(* IEC 61131-3 sources: traffic-lights/PLC_TrafficLights/Class/SafetyBaseFSoE (part 2) *)

  if WriteDOsUsed then
    for i := 0 to WriteDOsUsed-1 do
      SetDORunState(Handle:=aWritePDOs[i].Handle, NewState:=_BUS_IF_RUN_STATE_CONT_RUN);
    end_for;
  end_if;

  if usAnalogInputReadDOsUsed then
    for i := 0 to usAnalogInputReadDOsUsed-1 do
      SetDORunState(Handle:=aAnalogInputReadDOs[i].Handle, NewState:=_BUS_IF_RUN_STATE_CONT_RUN);
    end_for;
  end_if;

  if ReadFastUnsafeDOsUsed then
    for i := 0 to ReadFastUnsafeDOsUsed-1 do
      SetDORunState(Handle:=aFastUnsafeReadDOs[i].Handle, NewState:=_BUS_IF_RUN_STATE_CONT_RUN);
    end_for;
  end_if;

  if WriteFastUnsafeDOsUsed then
    for i := 0 to WriteFastUnsafeDOsUsed-1 do
      SetDORunState(Handle:=aFastUnsafeWriteDOs[i].Handle, NewState:=_BUS_IF_RUN_STATE_CONT_RUN);
    end_for;
  end_if;

END_FUNCTION

FUNCTION VIRTUAL SafetyBaseFSoE::StopDO
  VAR
    i : USINT;
  END_VAR

  // disable the DOs
  SetDORunState(Handle:=TempReadDO.Handle, NewState:=_BUS_IF_RUN_STATE_NO_RUN);

  SetDORunState(Handle:=TempWriteDO.Handle, NewState:=_BUS_IF_RUN_STATE_NO_RUN);

  if ReadDOsUsed then
    for i := 0 to ReadDOsUsed-1 do
      SetDORunState(Handle:=aReadPDOs[i].Handle, NewState:=_BUS_IF_RUN_STATE_NO_RUN);
    end_for;
  end_if;

  if WriteDOsUsed then
    for i := 0 to WriteDOsUsed-1 do
      SetDORunState(Handle:=aWritePDOs[i].Handle, NewState:=_BUS_IF_RUN_STATE_NO_RUN);
    end_for;
  end_if;

  if usAnalogInputReadDOsUsed then
    for i := 0 to usAnalogInputReadDOsUsed-1 do
      SetDORunState(Handle:=aAnalogInputReadDOs[i].Handle, NewState:=_BUS_IF_RUN_STATE_NO_RUN);
    end_for;
  end_if;

  if ReadFastUnsafeDOsUsed then
    for i := 0 to ReadFastUnsafeDOsUsed-1 do
      SetDORunState(Handle:=aFastUnsafeReadDOs[i].Handle, NewState:=_BUS_IF_RUN_STATE_NO_RUN);
    end_for;
  end_if;

  if WriteFastUnsafeDOsUsed then
    for i := 0 to WriteFastUnsafeDOsUsed-1 do
      SetDORunState(Handle:=aFastUnsafeWriteDOs[i].Handle, NewState:=_BUS_IF_RUN_STATE_NO_RUN);
    end_for;
  end_if;

END_FUNCTION

FUNCTION VIRTUAL SafetyBaseFSoE::InitBuffers
  VAR_OUTPUT
    sd_retval 	: DINT;
  END_VAR

  sd_retval := -1;

  //allocate memory for outgoing SDO (one SDO possible)
  p_SDOOutputBuffer$^void := ToStdLib.Malloc(size := SBF_SDO_MAX_LENGTH);

  if ( p_SDOOutputBuffer = NIL ) then
    SetSafetyState(NewState:=_MemAllocFailed);
    return;
  end_if;

  //allocate memory for incoming SDO list (number of SDO is dynamical)
  //following elements will be added dynamical

  //allocate list
  InputBufferAllocatedNo := SBF_SDO_BUFFER_ALLOC_BLOCK;
  p_SDOInputBuffer$^void := ToStdLib.Malloc(size := InputBufferAllocatedNo * SBF_SDO_MAX_LENGTH);

  if ( p_SDOInputBuffer = NIL ) then
    SetSafetyState(NewState:=_MemAllocFailed);
    return;
  end_if;

  //all buffers initialized
  sd_retval := 0;

END_FUNCTION

FUNCTION VIRTUAL SafetyBaseFSoE::GetSafetyNumber
  VAR_OUTPUT
    sd_retval 	: DINT;
  END_VAR
  VAR
    TempPathInfo  : PathInfoType;
    MyPara 	  : CmdStruct;
    MyResult	: results;
  END_VAR

  sd_retval := SDOStdRequ ( us_Command      := SBF_SDO_COMMAND_GET_SAFENBR
                          , p_us_RespData   := ( #SafetyNumber )$^USINT
                          , us_RespLength   := sizeof(SafetyNumber)
                          );

  if ( sd_retval <> 0 ) then
    if b_NoSafetyLogged = FALSE then
      b_NoSafetyLogged := TRUE;
      LogError("@01D8 (SafetyBaseFSoE::GetSafetyNumber) [SL] No Safety Number available!");
    end_if;
  elsif pConfigMem then
    // store safety number in config memory
    pConfigMem^$HDINT := SafetyNumber;
  end_if;

  sd_retval := SDOStdRequ ( us_Command      := SBF_SDO_COMMAND_GET_FW_VERSION
                          , p_us_RespData   := ( #sFirmwareVersion )$^USINT
                          , us_RespLength   := sizeof(FirmwareVersionType)
                          );

  if ( sd_retval = 0 ) then
    FirmwareVersion := sFirmwareVersion.RevMinor OR (sFirmwareVersion.RevMajor SHL 16);

    // Minor Versions starting with 9xxx mark Bootloader versions
    if (sFirmwareVersion.RevMinor >= 9000) & (sFirmwareVersion.RevMinor < 10000) then
      LogError("@01D9 (SafetyBaseFSoE::GetSafetyNumber) Bootloader version of safety firmware detected! Download a firmware or contact Sigmatek Support!");
    end_if;

    //Minor Versions higher than 338 mark versions which support the readout of the safety retry counters.
    if (sFirmwareVersion.RevMinor >= SBF_RETRY_COUNTER_AVAILABLE_MINOR_REV) & (sFirmwareVersion.RevMajor = SBF_RETRY_COUNTER_AVAILABLE_MAJOR_REV) then
      b_RetryCounterAvailable := TRUE;
    else
      b_RetryCounterAvailable := FALSE;
      //Call Method to set retrycounter servers of safety modules to -1
      SetRetryCounter();
    end_if;
  else
    SetSafetyState(NewState:=_ReadFWVerFailed);
    LogError("@01DA (SafetyBaseFSoE::GetSafetyNumber) No Firmware Version available!");
  end_if;

  InitPathInfo(#TempPathInfo);

  // add own safety number to routing table
  sd_retval := AddRoutingElement( ud_SafeNumber       := SafetyNumber
                                , ud_thisp            := this$UDINT
                                , pObject             := #TempPathInfo
                                );

  // give the manager more details about the module
  if pSafetyManagerThis then
    MyPara.uiCmd := CMD_SM_ADD_MODULE_INFO;
    MyPara.aPara[0] := THIS$DINT;
    MyPara.aPara[1] := SafetyNumber$DINT;
    MyPara.aPara[2] := FirmwareVersion$DINT;
    MyPara.aPara[3] := 16#FF; // fake FPGA_Version (only needed for CDIAS CPUs)
    MyPara.aPara[4] := to_DINT(p_ObjectPath^$USINT) + 1; // size of path (length + 1 for the length information)
    MyPara.aPara[5] := p_ObjectPath$DINT;
    pSafetyManagerThis^.NewInst(#MyPara, #MyResult);
  else
    LogError("@01DB (SafetyBaseFSoE::GetSafetyNumber) Couldn't find object of HwControl class, which is needed for safety time synchronisation!");
  end_if;

END_FUNCTION

FUNCTION SafetyBaseFSoE::SafetyBaseFSoE
  VAR_OUTPUT
    ret_code 	: ConfStates;
  END_VAR

#ifdef HWC_LogInit
  HWC_LogInit();
#endif

  //get interface for safety functions
  if ( OS_CILGET(INTERFACE_SAFETY, #pISafety)) then
    pISafety := NIL;

    LogError("@01DC (SafetyBaseFSoE::SafetyBaseFSoE) No Safety Interface found!");
  end_if;

  // initialize it with FALSE, if there is anything on local CDIAS it will change to TRUE
  b_SafetyOnLocalCDIAS := FALSE;

  // initialize module count with 0
  ModuleSyncNo := 0;

  ret_code := C_OK;

END_FUNCTION

#pragma warning(disable:0073);
FUNCTION VIRTUAL SafetyBaseFSoE::UpDateNotStd
  VAR_INPUT
    calloption 	: UDINT;
  END_VAR

END_FUNCTION
#pragma warning(default:0073);

FUNCTION VIRTUAL SafetyBaseFSoE::ReadSDOConfig
  VAR_INPUT
    p_SDORequestBuffer 	: ^SafetyBaseFSoE::SDORequReadConfig;
    p_SDOResponseBuffer 	: ^SafetyBaseFSoE::SDORespReadConfig;
    pModule 	: ^SafetyBaseFSoE::PathInfoType;
    pListHeader 	: ^SafetyBaseFSoE::PathInfoType;
  END_VAR
  VAR_OUTPUT
    sd_retval 	: DINT;
  END_VAR
  VAR
    ud_Address                    : UDINT;
    ud_ListLength_Address         : UDINT;
    ud_ListLength                 : UDINT;
    ud_TmpCnt                     : UDINT;
    i                             : UDINT;
    ud_ModulePathLen_Max          : UDINT;
    ud_ModulePathCompLen_Max      : UDINT;
    ud_ListHeaderPathLen_Max      : UDINT;
    ud_ListHeaderPathCompLen_Max  : UDINT;
    us_DataLength_Max             : USINT;
    ud_ListBaseAddress            : UDINT;
    ud_ListAddressMax             : UDINT;
    ud_CntUnsafeOutputs           : UDINT;
    ud_CntUnsafeInputs            : UDINT;
    ud_ActAddress                 : UDINT;  // actual offset in application memory (where to find the values in run mode)
    ud_UnsafeBDINT_Offset         : UDINT;  // actual offset in application memory (where to find the unsafe variables in run mode)
    ud_ActBlockType               : UDINT;
    ud_TmpAddress                 : UDINT;
    ud_TmpStrLen                  : UDINT;
    p_TmpBlockedData              : ^void;
    ud_ActStrLen                  : UDINT;
    us_BlockedTransferLength      : USINT;
    BoolOuts                      : UDINT;
    DintOuts                      : UDINT;
    TempModuleConfig              : t_ModuleCfg;
    pChar                         : ^CHAR;
    TempPath                      : ARRAY [0..99] OF USINT;
    PathOfThisCPU                 : ARRAY [0..99] OF USINT;
    GotOwnPath                    : BOOL;
    TempPdoConfig                 : t_PdoCfg;
    pBitMasks                     : ^BDINT;
    ActBitMask                    : BDINT;
    ud_skipLength                 : UDINT; //++pr
    b_CfgTypeV2                   : BOOL; // FALSE means there is no support of new time synchronisation/new general purpose register
    TmpCRC                        : HDINT;
    ud_ContainerBlockType         : UDINT;
    b_CfgTypeV3                   : BOOL;
    ud_ConfigLength               : UDINT;
    hd_DynParaVersion             : UDINT;
    DynamicParameterHeader        : t_DynamicParameterHeader;
    b_IsFSoE                      : BOOL;
    DynHeadSize                   : UDINT;
    AddressServiceDataSize        : UDINT;
    b_IprCodeLengthAvailable      : BOOL;  //TRUE, SCP211 is used
    ud_CntFastUnsafeOutputs       : UDINT;
    ud_CntFastUnsafeInputs        : UDINT;
    ud_FastUnsafe_Offset_In       : UDINT; // actual offset in application memory (where to find the unsafe variables in run mode)
    ud_FastUnsafe_Offset_Out      : UDINT; // actual offset in application memory (where to find the unsafe variables in run mode)
    ud_TmpLength                  : UDINT;

  END_VAR

  //minimum length of path: 2 bytes length, 1 byte domain info, 1 byte bus type and 1 byte port  => we use maximum so we don't have dynamic memory => don't fragment heap
  ud_ModulePathLen_Max          := 128;
  ud_ModulePathCompLen_Max      := 128;
  ud_ListHeaderPathLen_Max      := 128;
  ud_ListHeaderPathCompLen_Max  := 128;

  NewConfigType := ConfigState_NotInitialized;

  // reset flags before checking the config
  sFlexCon.FoundNodeInConfig := FALSE;
  sFlexCon.FoundHostInConfig := FALSE;
  b_IprCodeLengthAvailable        := FALSE;

  // also reset the servers
  if sFlexCon.pCommand & sFlexCon.pStateMachine & sFlexCon.pHostSafetyNumber then
    sFlexCon.pCommand^          := 0;
    sFlexCon.pStateMachine^     := 0;
    sFlexCon.pHostSafetyNumber^ := 0;
  end_if;

  //initialize header-data for request

  //calculate length without crc
  p_SDORequestBuffer^.StdHeader.Len := sizeof(SDORequReadConfig) - sizeof(SDOHeader.StdHeader.CRC);

  //type
  p_SDORequestBuffer^.StdHeader.Typ := SDO_STD;

  //command for reading config data
  p_SDORequestBuffer^.StdHeader.Cmd := SBF_SDO_COMMAND_READ;

  //read crc of whole config data

  //send request and receive data
  sd_retval := SDOReadCfgRequ ( p_SDORequestBuffer  := p_SDORequestBuffer
                              , p_SDOResponseBuffer := p_SDOResponseBuffer
                              , ud_Address          := SBF_SDO_ADDRESS_CONFIG_DATA + SBF_SDO_OFFSET_CONFIG_CRC_ALL
                              , us_Length           := 4
                              );

  //no response
  if ( sd_retval <> 0 ) then
    LogError("@01DD (SafetyBaseFSoE::ReadSDOConfig) Error reading CRC of config data.");
    return;
  end_if;

  // save crc and remember the time
  DesignerPrjConfigCRC := p_SDOResponseBuffer^.ud_Data;
  ud_LastCrcCheck := ops.tAbsolute;
  b_CheckCRC := TRUE;

  //read length of whole config data

  //send request and receive data
  sd_retval := SDOReadCfgRequ ( p_SDORequestBuffer  := p_SDORequestBuffer
                              , p_SDOResponseBuffer := p_SDOResponseBuffer
                              , ud_Address          := SBF_SDO_ADDRESS_CONFIG_DATA + SBF_SDO_OFFSET_CONFIG_LEN_ALL
                              , us_Length           := 4
                              );

  //no response
  if ( sd_retval <> 0 ) then
    LogError("@01DE (SafetyBaseFSoE::ReadSDOConfig) Error reading length of config data.");
    return;
  end_if;

  //no config data available
  if ( p_SDOResponseBuffer^.ud_Data = 16#FFFF_FFFF ) then
    LogError("@01DF (SafetyBaseFSoE::ReadSDOConfig) No config data available..");
    b_ReadConfigFailed := TRUE;
    return;
  end_if;

  ud_ConfigLength := p_SDOResponseBuffer^.ud_Data;

  // get BlockType
  //send request and receive data
  sd_retval := SDOReadCfgRequ ( p_SDORequestBuffer  := p_SDORequestBuffer
                              , p_SDOResponseBuffer := p_SDOResponseBuffer
                              , ud_Address          := SBF_SDO_ADDRESS_CONFIG_DATA + SBF_SDO_OFFSET_CONFIG_BLOCKTYPE
                              , us_Length           := 4
                              );
  //no response, error
  if ( sd_retval <> 0 ) then
    LogError("@01E0 (SafetyBaseFSoE::ReadSDOConfig) Error getting the block type of the header.");
    return;
  end_if;

  ud_ContainerBlockType := p_SDOResponseBuffer^.ud_Data;

  // check if it's a new version of the configuration
  if (ud_ContainerBlockType = SBF_BLKTYPE_CFG_CONTAINER_V3)       |
     (ud_ContainerBlockType = SBF_BLKTYPE_CFG_CONTAINER_V3_SLAVE)     |
     (ud_ContainerBlockType = SBF_BLKTYPE_CFG_CONTAINER_V3_SLAVE_OPTIONAL) then

    //read dynamic header length (how many data are attached to the header)

    //send request and receive data
    sd_retval := SDOReadCfgRequ ( p_SDORequestBuffer  := p_SDORequestBuffer
                                , p_SDOResponseBuffer := p_SDOResponseBuffer
                                , ud_Address          := SBF_SDO_ADDRESS_CONFIG_DATA + SBF_SDO_OFFSET_CONFIG_LEN_HEAD
                                , us_Length           := 4
                                );

    //no response
    if ( sd_retval <> 0 ) then
      LogError("@01E1 (SafetyBaseFSoE::ReadSDOConfig) Error reading length of dynamic header data.");
      return;
    end_if;

    // plausibility check for data length
    if p_SDOResponseBuffer^.ud_Data > 1000 then
      sd_retval := -1;
      LogError("@01E2 (SafetyBaseFSoE::ReadSDOConfig) Invalid length of dynamic header data.");
      return;
    end_if;

    // the length info contains: size of length info + size of time info + size of additional data

    //start address of first list: address of dynamic length + length according to length info
    ud_ListBaseAddress := SBF_SDO_ADDRESS_CONFIG_DATA + SBF_SDO_OFFSET_CONFIG_LEN_HEAD + p_SDOResponseBuffer^.ud_Data;

    DynHeadSize := p_SDOResponseBuffer^.ud_Data;

    // if we got at least 4 byte additional header data, it's the version of the dynamic parameters => read it
    if DynHeadSize >= 12 then
      //send request and receive data
      sd_retval := SDOReadCfgRequ ( p_SDORequestBuffer  := p_SDORequestBuffer
                                  , p_SDOResponseBuffer := p_SDOResponseBuffer
                                  , ud_Address          := SBF_SDO_ADDRESS_CONFIG_DATA + SBF_SDO_OFFSET_CONFIG_LEN_HEAD + 8
                                  , us_Length           := 4
                                  );

      //no response
      if ( sd_retval <> 0 ) then
        LogError("@01E3 (SafetyBaseFSoE::ReadSDOConfig) Error reading version of dynamic header data.");
        return;
      end_if;

      hd_DynParaVersion := p_SDOResponseBuffer^.ud_Data;
    else
      LogError("@01E4 (SafetyBaseFSoE::ReadSDOConfig) Data structure error in config! No bytes for the dynamic parameter version (according to length info).");
      return;
    end_if;

    // if we got at least 8 byte additional header data, the next 4 bytes are the flags => read it
    if DynHeadSize >= 16 then
      //send request and receive data
      sd_retval := SDOReadCfgRequ ( p_SDORequestBuffer  := p_SDORequestBuffer
                                  , p_SDOResponseBuffer := p_SDOResponseBuffer
                                  , ud_Address          := SBF_SDO_ADDRESS_CONFIG_DATA + SBF_SDO_OFFSET_CONFIG_LEN_HEAD + 12
                                  , us_Length           := 4
                                  );

      //no response
      if ( sd_retval <> 0 ) then
        LogError("@023D (SafetyBaseFSoE::ReadSDOConfig) Error reading flags of dynamic header data.");
        return;
      end_if;

      b_IsFSoE := (p_SDOResponseBuffer^.ud_Data AND 1) <> 0;

      // if we got the FSoE bit set => read the FSoE config
      if b_IsFSoE then
        GetFSoEConnectionInfos(p_SDORequestBuffer   := p_SDORequestBuffer
                             , p_SDOResponseBuffer  := p_SDOResponseBuffer
                             );
      end_if;

      if DynHeadSize >= 20 then
        //send request and receive data
        sd_retval := SDOReadCfgRequ ( p_SDORequestBuffer  := p_SDORequestBuffer
                                    , p_SDOResponseBuffer := p_SDOResponseBuffer
                                    , ud_Address          := SBF_SDO_ADDRESS_CONFIG_DATA + SBF_SDO_OFFSET_CONFIG_LEN_HEAD + 16
                                    , us_Length           := 4
                                    );

        //no response
        if ( sd_retval <> 0 ) then
          LogError("@023D (SafetyBaseFSoE::ReadSDOConfig) Error reading flags of dynamic header data.");
          return;
        end_if;

        b_IprCodeLengthAvailable := (p_SDOResponseBuffer^.ud_Data AND 1) <> 0;

        // if there are fast unsafe variables to read
        if uiPDOReadSizeFastUnsafeVar then

          //malloc FastUnsafe Output Buffer
          pFastUnsafeOutBuffer := ToStdLib.Malloc(size:=uiPDOReadSizeFastUnsafeVar);

          if pFastUnsafeOutBuffer = NIL then
            LogError("@0784 (SafetyBaseFSoE::ReadSDOConfig) Failed to allocate memory for outputbuffer.");
            return;
          else
            // init buffer
            _memset(dest:=pFastUnsafeOutBuffer, usByte:=0x00, cntr:=uiPDOReadSizeFastUnsafeVar);
          end_if;
        end_if;

        // if there are fast unsafe variables to write
        if uiPDOWriteSizeFastUnsafeVar then

          //malloc FastUnsafe Input Buffer
          pFastUnsafeInBuffer := ToStdLib.Malloc(size:=uiPDOWriteSizeFastUnsafeVar);

          if pFastUnsafeInBuffer = NIL then
            LogError("@0785 (SafetyBaseFSoE::ReadSDOConfig) Failed to allocate memory for inputbuffer.");
            return;
          else
            // init buffer
            _memset(dest:=pFastUnsafeInBuffer, usByte:=0x00, cntr:=uiPDOWriteSizeFastUnsafeVar);
          end_if;
        end_if;
      end_if;

    else
      LogError("@01E4 (SafetyBaseFSoE::ReadSDOConfig) Data structure error in config! No bytes for the dynamic parameter version (according to length info).");
      return;
    end_if;
  else
    // old version => no dynamic header, the first list starts where the dynamic header length would be

    //start address of first list: address of time info + size of time info
    ud_ListBaseAddress := SBF_SDO_ADDRESS_CONFIG_DATA + SBF_SDO_OFFSET_CONFIG_LEN_HEAD + sizeof(UDINT);
  end_if;

  GotOwnPath := FALSE;

  //highest address for config data
  ud_ListAddressMax := SDO_ADDRESS_CONFIG_DATA + SDO_OFFSET_CONFIG_LEN_ALL + ud_ConfigLength;

  //max. length of data to read with one request
  us_DataLength_Max := SBF_SDO_MAX_LENGTH - sizeof(SDORespReadConfig) + sizeof(SDORespReadConfig.ud_Data);

  while ( ud_ListBaseAddress < ud_ListAddressMax ) do

    //first read length of path in list-header

    //read path in list-header
    sd_retval := ReadModulePath ( p_SDORequestBuffer          := p_SDORequestBuffer
                                , p_SDOResponseBuffer         := p_SDOResponseBuffer
                                , p_ud_Address                := #ud_ListBaseAddress
                                , pModule                     := pListHeader
                                , p_ud_ModulePathLen_Max      := #ud_ListHeaderPathLen_Max
                                , p_ud_ModulePathCompLen_Max  := #ud_ListHeaderPathCompLen_Max
                                , us_SDOMaxDataSize           := us_DataLength_Max
                                );

    //no response, error
    if ( sd_retval <> 0 ) then
      LogError("@01E5 (SafetyBaseFSoE::ReadSDOConfig) Error reading module path out of config data.");
      return;
    end_if;

    // remember our own uncompressed path (first listheader path in the memory)
    if pListHeader^.p_us_Path & (GotOwnPath = FALSE) then
      GotOwnPath := TRUE;

      // remember the path
      _memcpy(ptr1:=#PathOfThisCPU[0], ptr2:=pListHeader^.p_us_Path, cntr:=(pListHeader^.p_us_Path$^UINT)^ + 2);
    end_if;

    //read length of download data in list-header (=LengthOverall) and save address
    //to calculate later the address of next list-header
    //address = last address + 4 byte (CRC)
    ud_ListLength_Address := ud_ListBaseAddress + 4;

    //send request and receive data
    sd_retval := SDOReadCfgRequ ( p_SDORequestBuffer  := p_SDORequestBuffer
                                , p_SDOResponseBuffer := p_SDOResponseBuffer
                                , ud_Address          := ud_ListLength_Address
                                , us_Length           := 4
                                );

    //no response
    if ( sd_retval <> 0 ) then
      LogError("@01E6 (SafetyBaseFSoE::ReadSDOConfig) Failed to read out the length of the download data within the configuration.");
      return;
    end_if;

    //save length of list
    ud_ListLength := p_SDOResponseBuffer^.ud_Data;

    //                                                   v
    //address of LengthOverall + 4 bytes (LengthOverall, BlockType, ModuleID)
    ud_Address := ud_ListLength_Address + 4;

    // get BlockType
    //send request and receive data
    sd_retval := SDOReadCfgRequ ( p_SDORequestBuffer  := p_SDORequestBuffer
                                , p_SDOResponseBuffer := p_SDOResponseBuffer
                                , ud_Address          := ud_Address
                                , us_Length           := 4
                                );
    //no response, error
    if ( sd_retval <> 0 ) then
      LogError("@01E7 (SafetyBaseFSoE::ReadSDOConfig) Error getting the block type.");
      return;
    end_if;

    ud_ActBlockType := p_SDOResponseBuffer^.ud_Data;

    case ud_ActBlockType of
//**********************************************************************************************************************************************************
      SBF_BLKTYPE_CFG_CPU,
      SBF_BLKTYPE_CFG_CPU_OPTIONAL , // if we don't need data from an external cpu
      SBF_BLKTYPE_CFG_MASTER_CPU:
        //add other CPUs to routing table

        // if there is a valid module path
        if pListHeader^.p_us_Path <> NIL then
          //add module to routing tabs
          sd_retval := AddModuleToRoutingTabs ( pModule       := pListHeader
                                              , pListHeader   := pListHeader
                                              , b_IsOptional  := (ud_ActBlockType = SBF_BLKTYPE_CFG_CPU_OPTIONAL)
                                              );

          if (sd_retval <> 0 ) then
            if ( SafetyState <> _ModFromCfgNotFound ) then
              LogError("@01E8 (SafetyBaseFSoE::ReadSDOConfig) Failed to add cpu module to routing tabs.");
              return;
            end_if;
          end_if;

          TempModuleConfig.Info := 0;
          TempModuleConfig.DestCRCNo := 0;
          TempModuleConfig.pDestCRCs := NIL;
          TempModuleConfig.PdoOutLen := 0;

          TempModuleConfig.Info.IsOptional  := (ud_ActBlockType = SBF_BLKTYPE_CFG_CPU_OPTIONAL);
          TempModuleConfig.InterfaceCRC     := 0;

          // Remember the path (uncompressed and compressed)
          TempModuleConfig.PathLen := pListHeader^.p_us_Path^$UINT + 2;
          TempModuleConfig.pPath := pListHeader^.p_us_Path;

          TempModuleConfig.CompPathLen := pListHeader^.ui_PathCompLen;
          TempModuleConfig.pCompPath := pListHeader^.p_us_PathComp;

          // if it's our own path, remember the safety number
          if (PathOfThisCPU[0]$UINT = (pListHeader^.p_us_Path$^UINT)^) & (ToStdLib.MemCmp(#PathOfThisCPU[0], pListHeader^.p_us_Path, PathOfThisCPU[0]$UINT + 2) = 0) then
            TempModuleConfig.SafetyNbr := SafetyNumber;
            //safe config of scp modul (own path)
            SafeActModuleConfig(TempModuleConfig);
          else
            TempModuleConfig.SafetyNbr := 0;
          end_if;

          // only when there is a manager
          if pSafetyManagerThis then
            AddModuleToCfg(TempModuleConfig);
          end_if;
        end_if;

//**********************************************************************************************************************************************************
      SBF_BLKTYPE_CFG_SLAVE_COMPR,
      SBF_BLKTYPE_CFG_SLAVE_COMPR_OPTIONAL: //Blocktyp der über die komprimierte Gesamtkonfiguration einer Slave-CPU gegeben wird
        //add other CPUs to routing table

        // if there is a valid module path
        if pListHeader^.p_us_Path <> NIL then
          //add module to routing tabs
          sd_retval := AddModuleToRoutingTabs ( pModule       := pListHeader
                                              , pListHeader   := pListHeader
                                              , b_IsOptional  := (ud_ActBlockType = SBF_BLKTYPE_CFG_SLAVE_COMPR_OPTIONAL)
                                              );

          if (sd_retval <> 0 ) then
            if ( SafetyState <> _ModFromCfgNotFound ) then
              LogError("@0270 (SafetyBaseFSoE::ReadSDOConfig) Slave: Failed to add cpu module to routing tabs.");
              return;
            end_if;
          end_if;

          // we skip the config till we get to the interface information of this slave (if it's the source of an interface frame we have to remember it)

          //address of LengthOverall + 3 * 4 bytes (LengthOverall, BlockType, ModuleID) => now the address points to FUB offset
          ud_Address := ud_ListLength_Address + 12;

          //skip FUB offset
          ud_Address += 4;

          // get no of FUB´s
          //send request and receive data
          sd_retval := SDOReadCfgRequ ( p_SDORequestBuffer  := p_SDORequestBuffer
                                      , p_SDOResponseBuffer := p_SDOResponseBuffer
                                      , ud_Address          := ud_Address
                                      , us_Length           := 4
                                      );
          //no response, error
          if ( sd_retval <> 0 ) then
            LogError("@01E9 (SafetyBaseFSoE::ReadSDOConfig) Slave: Error getting the FUB number.");
            return;
          end_if;

          ud_TmpCnt := p_SDOResponseBuffer^.ud_Data;

          // skip no of FUB´s and FUB´s
          ud_Address += (4 + (ud_TmpCnt * 4));

          // get length of path
          //send request and receive data
          sd_retval := SDOReadCfgRequ ( p_SDORequestBuffer  := p_SDORequestBuffer
                                      , p_SDOResponseBuffer := p_SDOResponseBuffer
                                      , ud_Address          := ud_Address
                                      , us_Length           := 4
                                      );
          //no response, error
          if ( sd_retval <> 0 ) then
            LogError("@01EA (SafetyBaseFSoE::ReadSDOConfig) Slave: Error getting the path length.");
            return;
          end_if;

          ud_TmpCnt := p_SDOResponseBuffer^.ud_Data;

          // skip length of path and the path
          ud_Address += (4 + ud_TmpCnt);

          // get length of comp path
          //send request and receive data
          sd_retval := SDOReadCfgRequ ( p_SDORequestBuffer  := p_SDORequestBuffer
                                      , p_SDOResponseBuffer := p_SDOResponseBuffer
                                      , ud_Address          := ud_Address
                                      , us_Length           := 4
                                      );
          //no response, error
          if ( sd_retval <> 0 ) then
            LogError("@01EB (SafetyBaseFSoE::ReadSDOConfig) Slave: Error getting the comp path length.");
            return;
          end_if;

          ud_TmpCnt := p_SDOResponseBuffer^.ud_Data;

          // skip length of comp path and the comp path
          ud_Address += (4 + ud_TmpCnt);

          // skip CRC and LengthOverall to get to the Blocktyp (Modul-Downloaddaten)
          ud_Address += 8;

          // get the block type
          //send request and receive data
          sd_retval := SDOReadCfgRequ ( p_SDORequestBuffer  := p_SDORequestBuffer
                                      , p_SDOResponseBuffer := p_SDOResponseBuffer
                                      , ud_Address          := ud_Address
                                      , us_Length           := 4
                                      );
          //no response, error
          if ( sd_retval <> 0 ) then
            LogError("@01EC (SafetyBaseFSoE::ReadSDOConfig) Slave: Error getting the block type of a slave config.");
            return;
          end_if;

          ud_TmpCnt := p_SDOResponseBuffer^.ud_Data;

          // check if it's a new version of the configuration
          if (ud_TmpCnt = SBF_BLKTYPE_CFG_CONTAINER_V3)       |
             (ud_TmpCnt = SBF_BLKTYPE_CFG_CONTAINER_V3_SLAVE)     |
             (ud_TmpCnt = SBF_BLKTYPE_CFG_CONTAINER_V3_SLAVE_OPTIONAL) then

            // skip blocktype to get to the dynamic header length (how many data are attached to the header)
            ud_Address += 4;

            //send request and receive data
            sd_retval := SDOReadCfgRequ ( p_SDORequestBuffer  := p_SDORequestBuffer
                                        , p_SDOResponseBuffer := p_SDOResponseBuffer
                                        , ud_Address          := ud_Address
                                        , us_Length           := 4
                                        );

            //no response
            if ( sd_retval <> 0 ) then
              LogError("@01ED (SafetyBaseFSoE::ReadSDOConfig) Error reading length of dynamic header data of a slave config.");
              return;
            end_if;

            // plausibility check for data length
            if p_SDOResponseBuffer^.ud_Data > 1000 then
              sd_retval := -1;
              LogError("@01EE (SafetyBaseFSoE::ReadSDOConfig) Invalid length of dynamic header data of a slave config.");
              return;
            end_if;

            // the length info contains: size of length info + size of time info + size of additional data

            // skip the additional data to get to the path length
            ud_Address += p_SDOResponseBuffer^.ud_Data;
          else
            // old version => no dynamic header, so we skip only blocktype and time info
            ud_Address += 8;
          end_if;

          // get the path length
          //send request and receive data
          sd_retval := SDOReadCfgRequ ( p_SDORequestBuffer  := p_SDORequestBuffer
                                      , p_SDOResponseBuffer := p_SDOResponseBuffer
                                      , ud_Address          := ud_Address
                                      , us_Length           := 4
                                      );
          //no response, error
          if ( sd_retval <> 0 ) then
            LogError("@01EA (SafetyBaseFSoE::ReadSDOConfig) Slave: Error getting the path length.");
            return;
          end_if;

          ud_TmpCnt := p_SDOResponseBuffer^.ud_Data;

          // skip length of path and the path
          ud_Address += (4 + ud_TmpCnt);

          // get length of comp path
          //send request and receive data
          sd_retval := SDOReadCfgRequ ( p_SDORequestBuffer  := p_SDORequestBuffer
                                      , p_SDOResponseBuffer := p_SDOResponseBuffer
                                      , ud_Address          := ud_Address
                                      , us_Length           := 4
                                      );
          //no response, error
          if ( sd_retval <> 0 ) then
            LogError("@01EB (SafetyBaseFSoE::ReadSDOConfig) Slave: Error getting the comp path length.");
            return;
          end_if;

          ud_TmpCnt := p_SDOResponseBuffer^.ud_Data;

          // skip length of comp path and the comp path
          ud_Address += (4 + ud_TmpCnt);

          // skip CRC, LengthOverall, Blocktyp (Modul-Downloaddaten), ModuleID
          ud_Address += 16;

          // get the InterfaceCRC
          //send request and receive data
          sd_retval := SDOReadCfgRequ ( p_SDORequestBuffer  := p_SDORequestBuffer
                                      , p_SDOResponseBuffer := p_SDOResponseBuffer
                                      , ud_Address          := ud_Address
                                      , us_Length           := 4
                                      );
          //no response, error
          if ( sd_retval <> 0 ) then
            LogError("@01EF (SafetyBaseFSoE::ReadSDOConfig) Slave: Error getting the Inteface-CRC.");
            return;
          end_if;

          TmpCRC := p_SDOResponseBuffer^.ud_Data;

          //add slave information to config
          AddSlaveToCfg ( pModule       := pListHeader
                        , b_IsOptional  := (ud_ActBlockType = SBF_BLKTYPE_CFG_SLAVE_COMPR_OPTIONAL)
                        , b_IsInterface := (TmpCRC <> 0)
                        , InterfaceCRC  := TmpCRC
                        );

        end_if;

//**********************************************************************************************************************************************************
      SBF_BLKTYPE_CFG_REV: // revision

        // check if the list is long enough for a String (more bytes than just the header)
        if ud_ListLength > 12 then

          //address of LengthOverall + 3 * 4 bytes (LengthOverall, BlockType, ModuleID) => now the address points to the revision string
          ud_Address := ud_ListLength_Address + 12;

          //read out the string (length = LengthOverall - length header)

          // get memory for the string
          if pPrjNameStr = NIL then
            PrjNameMemLen := ud_ListLength$USINT - 12;
            pPrjNameStr$^void := ToStdLib.Malloc(size := PrjNameMemLen + 1);
          else
            if PrjNameMemLen <> (ud_ListLength$USINT - 12) then
              PrjNameMemLen := ud_ListLength$USINT - 12;
              pPrjNameStr$^void := ToStdLib.ReAlloc(mptr:=pPrjNameStr, newsize:=PrjNameMemLen + 1);
            end_if;
          end_if;

          // check if we got a memory
          if pPrjNameStr then

            _memset(dest:=pPrjNameStr, usByte:=0, cntr:=PrjNameMemLen+1);

            ud_ActStrLen := ud_TmpStrLen := PrjNameMemLen;
            ud_TmpAddress := ud_Address;

            IF p_BlockedTransferMemory = NIL THEN
              sd_retval := -100;
              SetSafetyState(NewState:=_MemAllocFailed);
              RETURN;
            END_IF;

            IF ud_BlockedTransferMemorySize < (ud_TmpStrLen + 1) THEN
              p_BlockedTransferMemory := ToStdLib.ReAlloc(mptr:=p_BlockedTransferMemory, newsize:=GetNewMemSize(ud_TmpStrLen + 1));
              IF p_BlockedTransferMemory = NIL THEN
                ud_BlockedTransferMemorySize := 0;
                sd_retval := -100;
                SetSafetyState(NewState:=_MemAllocFailed);
                RETURN;
              ELSE
                ud_BlockedTransferMemorySize := GetNewMemSize(ud_TmpStrLen + 1);
              END_IF;
            END_IF;

            ToStdLib.MemSet(dest:=p_BlockedTransferMemory, value:=0, size:=ud_BlockedTransferMemorySize);

            p_TmpBlockedData := p_BlockedTransferMemory;

            us_BlockedTransferLength := BlockedTransferLength(ud_Datalength:=ud_TmpStrLen, us_MaxBlocklength:=60);

            while us_BlockedTransferLength do

              // get name
              sd_retval := SDOReadCfgRequ ( p_SDORequestBuffer  := p_SDORequestBuffer
                                          , p_SDOResponseBuffer := p_SDOResponseBuffer
                                          , ud_Address          := ud_TmpAddress
                                          , us_Length           := us_BlockedTransferLength
                                          , b_UseCache          := us_BlockedTransferLength < us_DataLength_Max
                                          );
              //no response
              if ( sd_retval <> 0 ) then
                LogError("@01F0 (SafetyBaseFSoE::ReadSDOConfig) Reading Revision failed.");
                return;
              end_if;

              ToStdLib.MemCpy(dest:=p_TmpBlockedData,
                               source:=#p_SDOResponseBuffer^.ud_Data,
                               size:=us_BlockedTransferLength);

              p_TmpBlockedData += us_BlockedTransferLength;
              ud_TmpAddress += us_BlockedTransferLength;
              ud_TmpStrLen -= us_BlockedTransferLength;

              us_BlockedTransferLength := BlockedTransferLength(ud_Datalength:=ud_TmpStrLen, us_MaxBlocklength:=60);

            end_while;

            ToStdLib.MemCpy(dest:=pPrjNameStr,
                             source:=p_BlockedTransferMemory,
                             size:=PrjNameMemLen+1);

            b_GotNewRevision := TRUE;

            // string is formed by: project name {TAB} project revision   => search for the tab
            pPrjRevStr := pPrjNameStr; // initialize pointer, because maybe there is no content in the projectname
            pChar := pPrjNameStr;
            while pChar^ do
              // check for tab sign
              if pChar^ = 9 then
                // at the next character our revision starts
                pPrjRevStr := pChar + sizeof(CHAR);

                // we change the tab to a string termination
                pChar^ := 0;

                // save the length of the name and the length of the project revision
                PrjNameStrLen := pChar$UDINT - pPrjNameStr$UDINT;
                PrjRevStrLen := PrjNameMemLen - PrjNameStrLen - sizeof(CHAR);
                exit;
              end_if;

              pChar += sizeof(CHAR);
            end_while;

            ShowProjectRevision();
          end_if;
        end_if;

//**********************************************************************************************************************************************************
      SBF_BLKTYPE_CFG_CRC: // CRC from Safety Application and HW-Tree

        // check if the list is long enough for a String (more bytes than just the header)
        if ud_ListLength > 12 then

          //address of LengthOverall + 3 * 4 bytes (LengthOverall, BlockType, ModuleID) => now the address points to the CRC values
          ud_Address := ud_ListLength_Address + 12;

          //read out the CRCs (length = 2 * 4 bytes)

          //send request and receive data
          sd_retval := SDOReadCfgRequ ( p_SDORequestBuffer  := p_SDORequestBuffer
                                      , p_SDOResponseBuffer := p_SDOResponseBuffer
                                      , ud_Address          := ud_Address
                                      , us_Length           := 2*sizeof(HDINT)
                                      );

          //no response
          if ( sd_retval <> 0 ) then
            LogError("@0797 (SafetyBaseFSoE::ReadSDOConfig) Reading CRC info of the safety designer project failed.");
            return;
          end_if;

          CRCInfo := p_SDOResponseBuffer^.ud_Data$t_CRCInfo;

          ApplCRC := CRCInfo.ApplCRC;
          HwCRC   := CRCInfo.HwCRC;
        end_if;

//**********************************************************************************************************************************************************
      SBF_BLKTYPE_CFG_INTERFACE,
      SBF_BLKTYPE_CFG_INTERFACE_OPTIONAL: // interface frame

        TempPdoConfig.Info := 0;

        //address of LengthOverall + 3 * 4 bytes (LengthOverall, BlockType, Module ID) => points to interface CRC
        ud_Address := ud_ListLength_Address + 12;

//*****************************************************************************
//**   INTERFACE CRC                                                         **
//*****************************************************************************

        //send request and receive data
        sd_retval := SDOReadCfgRequ ( p_SDORequestBuffer  := p_SDORequestBuffer
                                    , p_SDOResponseBuffer := p_SDOResponseBuffer
                                    , ud_Address          := ud_Address
                                    , us_Length           := 4
                                    );

        //no response
        if ( sd_retval <> 0 ) then
          LogError("@01F1 (SafetyBaseFSoE::ReadSDOConfig) Interface: Reading interface CRC of interface frame block failed.");
          return;
        end_if;

        TempPdoConfig.InterfaceCRC := p_SDOResponseBuffer^.ud_Data;

        // skip interface crc
        ud_Address += 4;

//*****************************************************************************
//**   LENGTH OF TOPOLOGY PATH OF INTERFACE FRAME                            **
//*****************************************************************************

        //send request and receive data
        sd_retval := SDOReadCfgRequ ( p_SDORequestBuffer  := p_SDORequestBuffer
                                    , p_SDOResponseBuffer := p_SDOResponseBuffer
                                    , ud_Address          := ud_Address
                                    , us_Length           := 4
                                    );

        //no response
        if ( sd_retval <> 0 ) then
          LogError("@01F2 (SafetyBaseFSoE::ReadSDOConfig) Interface: Reading length of topology path of interface frame block failed.");
          return;
        end_if;

        // skip path length
        ud_Address += 4;

        us_BlockedTransferLength := p_SDOResponseBuffer^.ud_Data$USINT;

//*****************************************************************************
//**   TOPOLOGY PATH OF INTERFACE FRAME                                      **
//*****************************************************************************

        //send request and receive data
        sd_retval := SDOReadCfgRequ ( p_SDORequestBuffer  := p_SDORequestBuffer
                                    , p_SDOResponseBuffer := p_SDOResponseBuffer
                                    , ud_Address          := ud_Address
                                    , us_Length           := us_BlockedTransferLength
                                    , b_UseCache          := us_BlockedTransferLength < us_DataLength_Max
                                    );

        //no response
        if ( sd_retval <> 0 ) then
          LogError("@01F3 (SafetyBaseFSoE::ReadSDOConfig) Interface: Reading topology path of interface frame block failed.");
          return;
        end_if;

        // remember the destination path
        _memcpy(ptr1:=#TempPath[0], ptr2:=#p_SDOResponseBuffer^.ud_Data, cntr:=us_BlockedTransferLength);

        // this is the source of the interface frame
        TempPdoConfig.SourcePathLen := TempPath[0]$UINT + 2;
        TempPdoConfig.pSourcePath   := #TempPath[0];

        // skip path
        ud_Address += us_BlockedTransferLength;

//*****************************************************************************
//**   LENGTH OF COMPRESSED TOPOLOGY PATH OF INTERFACE FRAME                 **
//*****************************************************************************

        //send request and receive data
        sd_retval := SDOReadCfgRequ ( p_SDORequestBuffer  := p_SDORequestBuffer
                                    , p_SDOResponseBuffer := p_SDOResponseBuffer
                                    , ud_Address          := ud_Address
                                    , us_Length           := 4
                                    );

        //no response
        if ( sd_retval <> 0 ) then
          LogError("@01F4 (SafetyBaseFSoE::ReadSDOConfig) Interface: Reading length of compressed topology path of interface frame block failed.");
          return;
        end_if;

        // skip path length
        ud_Address += 4;

        us_BlockedTransferLength := p_SDOResponseBuffer^.ud_Data$USINT;

//*****************************************************************************
//**   COMPRESSED TOPOLOGY PATH OF INTERFACE FRAME                           **
//*****************************************************************************

        //send request and receive data
        sd_retval := SDOReadCfgRequ ( p_SDORequestBuffer  := p_SDORequestBuffer
                                    , p_SDOResponseBuffer := p_SDOResponseBuffer
                                    , ud_Address          := ud_Address
                                    , us_Length           := us_BlockedTransferLength
                                    , b_UseCache          := us_BlockedTransferLength < us_DataLength_Max
                                    );

        //no response
        if ( sd_retval <> 0 ) then
          LogError("@01F5 (SafetyBaseFSoE::ReadSDOConfig) Interface: Reading compressed topology path of interface frame block failed.");
          return;
        end_if;

        // if it's an IP address => we need the compressed path for the source
        if p_SDOResponseBuffer^.ud_Data$USINT = 6 then
          // we may need this later (e.g. if it's an IP address)
          _memcpy(ptr1:=#TempPath[0], ptr2:=#p_SDOResponseBuffer^.ud_Data, cntr:=us_BlockedTransferLength);

          // this is the source of the interface frame
          TempPdoConfig.SourcePathLen := us_BlockedTransferLength;
          TempPdoConfig.Info.SrcPathIsCompressed := TRUE;

          if ((#p_SDOResponseBuffer^.ud_Data + 5)^$HDINT AND 16#00FFFFFF) = 0 then
            // special IP: (0.0.0.x)
            TempPdoConfig.Info.SrcPathIsCompressed := FALSE;  // Not valid IP
          end_if;
        end_if;

        // skip path and maximum cycle time
        ud_Address += us_BlockedTransferLength + 4;

  // here starts the data area (before we read only the list header

//*****************************************************************************
//**   INTERFACE CRC                                                         **
//*****************************************************************************

        //send request and receive data
        sd_retval := SDOReadCfgRequ ( p_SDORequestBuffer  := p_SDORequestBuffer
                                    , p_SDOResponseBuffer := p_SDOResponseBuffer
                                    , ud_Address          := ud_Address
                                    , us_Length           := 4
                                    );

        //no response
        if ( sd_retval <> 0 ) then
          LogError("@01F6 (SafetyBaseFSoE::ReadSDOConfig) Interface: Reading CRC of interface frame block failed.");
          return;
        end_if;

        TempPdoConfig.InterfaceCRC := p_SDOResponseBuffer^.ud_Data;

        // skip interface CRC
        ud_Address += 4;

//*****************************************************************************
//**   NUMBER OF BOOL INTERFACE VARIABLES IN THE PDO                         **
//*****************************************************************************

        //send request and receive data
        sd_retval := SDOReadCfgRequ ( p_SDORequestBuffer  := p_SDORequestBuffer
                                    , p_SDOResponseBuffer := p_SDOResponseBuffer
                                    , ud_Address          := ud_Address
                                    , us_Length           := 4
                                    );

        //no response
        if ( sd_retval <> 0 ) then
          LogError("@01F7 (SafetyBaseFSoE::ReadSDOConfig) Interface: Reading number of bool variables in the interface frame failed.");
          return;
        end_if;

        BoolOuts := p_SDOResponseBuffer^.ud_Data;

        // skip bool variables
        ud_Address += 4;

//*****************************************************************************
//**   NUMBER OF DINT INTERFACE VARIABLES IN THE PDO                         **
//*****************************************************************************

        //send request and receive data
        sd_retval := SDOReadCfgRequ ( p_SDORequestBuffer  := p_SDORequestBuffer
                                    , p_SDOResponseBuffer := p_SDOResponseBuffer
                                    , ud_Address          := ud_Address
                                    , us_Length           := 4
                                    );

        //no response
        if ( sd_retval <> 0 ) then
          LogError("@01F8 (SafetyBaseFSoE::ReadSDOConfig) Interface: Reading number of dint variables in the interface frame failed.");
          return;
        end_if;

        // skip dint variables
        ud_Address += 4;

        DintOuts := p_SDOResponseBuffer^.ud_Data;

        // if there are interface variables
        if BoolOuts | DintOuts then
          // calculate the length of the interface frame
          TempPdoConfig.PdoLen := CalcPDOLength(BoolOuts, DintOuts);

          // and the destination
          TempPdoConfig.DestPathLen   := PathOfThisCPU[0]$UINT + 2;
          TempPdoConfig.pDestPath     := #PathOfThisCPU[0];

          TempPdoConfig.Info.IsInterfacePDO := TRUE;
          TempPdoConfig.Info.IsOptional := (ud_ActBlockType = SBF_BLKTYPE_CFG_INTERFACE_OPTIONAL);

          // add the interface PDO to the list
          AddPdoToCfg(TempPdoConfig);
        else
          LogError("@01F9 (SafetyBaseFSoE::ReadSDOConfig) Interface: No interface variables found in interface blocktype.");
          return;
        end_if;

//**********************************************************************************************************************************************************
      SBF_BLKTYPE_CFG_MODULE_WITHOUT_CFG,
      SBF_BLKTYPE_CFG_MODULE_WITHOUT_CFG_OPT:      // module configurations
        TempModuleConfig.Info := 0;
        TempModuleConfig.DestCRCNo := 0;
        TempModuleConfig.pDestCRCs := NIL;
        case ud_ActBlockType of
          SBF_BLKTYPE_CFG_MODULE_WITHOUT_CFG_OPT:
            TempModuleConfig.Info.IsOptional := TRUE;
          else
            TempModuleConfig.Info.IsOptional := FALSE;
        end_case;

        BoolOuts := 0;
        DintOuts := 0;

        // Remember the path (uncompressed and compressed)
        TempModuleConfig.PathLen := pListHeader^.p_us_Path^$UINT + 2;
        TempModuleConfig.pPath := pListHeader^.p_us_Path;

        TempModuleConfig.CompPathLen := pListHeader^.ui_PathCompLen;
        TempModuleConfig.pCompPath := pListHeader^.p_us_PathComp;

        //add module to routing tabs
        sd_retval := AddModuleToRoutingTabs ( pModule       := pListHeader
                                            , pListHeader   := pListHeader
                                            , b_IsOptional  := TempModuleConfig.Info.IsOptional
                                            );

        if (sd_retval <> 0 ) then
          if ( SafetyState <> _ModFromCfgNotFound ) then
            LogError("@020D (SafetyBaseFSoE::ReadSDOConfig) Failed to add safe input module to routing tabs.");
            return;
          end_if;
        end_if;

//*****************************************************************************
//**   LIST HEADER                                                           **
//*****************************************************************************
//   Offset  Größe	Beschreibung
//    0x00	4 Byte	CRC32
//    0x04	4 Byte	Länge der Konfiguration (inkl. Längenfeld)
//    0x08	4 Byte	Block-Typ (nicht optional: 0x00000029; optional: 0x40000029)
//    0x0C	4 Byte	Modul-ID
//    0x10	4 Byte	Version der Konfiguration (0x00000000)
//*****************************************************************************

        //address of LengthOverall + 4 * 4 bytes (LengthOverall, BlockType, ModuleID, VersionConfig)
        ud_Address := ud_ListLength_Address + 16;

//*****************************************************************************
//    FSoE Konfiguration
//*****************************************************************************
//    0x14	4 Byte	Anzahl an FSoE-Verbindungen (0x00000001)
//*****************************************************************************
//    FSoE Konfiguration * Anzahl an FSoE-Verbindungen
//*****************************************************************************
//    0x18	4 Byte	Länge der FSoE-Konfiguration
//    0x1C	4 Byte	Flags (0x00000000)
//    0x20	2 Byte	Größe der sicheren Ausgänge in Byte
//    0x22	2 Byte	Größe der sicheren Eingänge in Byte
//    0x24	2 Byte	FSoE Slaveadresse
//    0x26	2 Byte	reserviert
//*****************************************************************************

        // skip entrys to read fsoe slave address
        ud_Address += 16;

        //send request and receive data
        sd_retval := SDOReadCfgRequ ( p_SDORequestBuffer  := p_SDORequestBuffer
                                    , p_SDOResponseBuffer := p_SDOResponseBuffer
                                    , ud_Address          := ud_Address
                                    , us_Length           := 4
                                    );

        //no response
        if ( sd_retval <> 0 ) then
          LogError("@01F6 (SafetyBaseFSoE::ReadSDOConfig) Reading interface CRC of interface frame block failed.");
          return;
        end_if;

        // only when there is a manager
        if pSafetyManagerThis then
          AddModuleToCfg(TempModuleConfig);
        end_if;

//**********************************************************************************************************************************************************
      SBF_BLKTYPE_CFG_MODULE,
      SBF_BLKTYPE_CFG_MODULE_V2,
      SBF_BLKTYPE_CFG_MODULE_OPTIONAL,
      SBF_BLKTYPE_CFG_CONTAINER_SLAVE,
      SBF_BLKTYPE_CFG_CONTAINER_SLAVE_OPTIONAL,
      SBF_BLKTYPE_CFG_MODULE_V3,
      SBF_BLKTYPE_CFG_MODULE_V3_OPTIONAL,
      SBF_BLKTYPE_CFG_CONTAINER_V3_SLAVE,
      SBF_BLKTYPE_CFG_CONTAINER_V3_SLAVE_OPTIONAL:      // module configurations
        TempModuleConfig.Info := 0;
        TempModuleConfig.DestCRCNo := 0;
        TempModuleConfig.pDestCRCs := NIL;
        case ud_ActBlockType of
          SBF_BLKTYPE_CFG_MODULE_OPTIONAL,
          SBF_BLKTYPE_CFG_CONTAINER_SLAVE_OPTIONAL,
          SBF_BLKTYPE_CFG_MODULE_V3_OPTIONAL,
          SBF_BLKTYPE_CFG_CONTAINER_V3_SLAVE_OPTIONAL:
            TempModuleConfig.Info.IsOptional := TRUE;
          else
            TempModuleConfig.Info.IsOptional := FALSE;
        end_case;

        b_CfgTypeV2 := (ud_ActBlockType <> SBF_BLKTYPE_CFG_MODULE);

        // check if it's a V3 config, because the structure of the IO List is different
        if (ud_ActBlockType = SBF_BLKTYPE_CFG_MODULE_V3) |
           (ud_ActBlockType = SBF_BLKTYPE_CFG_MODULE_V3_OPTIONAL) |
           (ud_ActBlockType = SBF_BLKTYPE_CFG_CONTAINER_V3_SLAVE) |
           (ud_ActBlockType = SBF_BLKTYPE_CFG_CONTAINER_V3_SLAVE_OPTIONAL) then
          b_CfgTypeV3 := TRUE;
        else
          b_CfgTypeV3 := FALSE;
        end_if;

        // if it's our own path, remember the type of module configuration
        if (PathOfThisCPU[0]$UINT = (pListHeader^.p_us_Path$^UINT)^) & (ToStdLib.MemCmp(#PathOfThisCPU[0], pListHeader^.p_us_Path, PathOfThisCPU[0]$UINT + 2) = 0) then
          // if config is already "old" dont change to "new". (can be set by block SBF_BLKTYPE_OLD_MODE_FLAG)
          if NewConfigType <> ConfigState_Old then
            NewConfigType := (b_CfgTypeV2$USINT + 1)$t_ConfigStateType;
          end_if;
        end_if;

        BoolOuts := 0;
        DintOuts := 0;

        // Remember the path (uncompressed and compressed)
        TempModuleConfig.PathLen := pListHeader^.p_us_Path^$UINT + 2;
        TempModuleConfig.pPath := pListHeader^.p_us_Path;

        TempModuleConfig.CompPathLen := pListHeader^.ui_PathCompLen;
        TempModuleConfig.pCompPath := pListHeader^.p_us_PathComp;

//*****************************************************************************
//**   LIST HEADER                                                           **
//*****************************************************************************

        //address of LengthOverall + 3 * 4 bytes (LengthOverall, BlockType, ModuleID)
        ud_Address := ud_ListLength_Address + 12;

        // only available at new modules
        if b_CfgTypeV2 then

//*****************************************************************************
//**   INTERFACE CRC                                                         **
//*****************************************************************************

          //send request and receive data
          sd_retval := SDOReadCfgRequ ( p_SDORequestBuffer  := p_SDORequestBuffer
                                      , p_SDOResponseBuffer := p_SDOResponseBuffer
                                      , ud_Address          := ud_Address
                                      , us_Length           := 4
                                      );

          //no response
          if ( sd_retval <> 0 ) then
            LogError("@01F6 (SafetyBaseFSoE::ReadSDOConfig) Reading interface CRC of interface frame block failed.");
            return;
          end_if;

          TempPdoConfig.InterfaceCRC := p_SDOResponseBuffer^.ud_Data;

          // skip interface crc
          ud_Address += 4;

//*****************************************************************************
//**   LENGTH OF TOPOLOGY PATH OF INTERFACE FRAME                            **
//*****************************************************************************

          //send request and receive data
          sd_retval := SDOReadCfgRequ ( p_SDORequestBuffer  := p_SDORequestBuffer
                                      , p_SDOResponseBuffer := p_SDOResponseBuffer
                                      , ud_Address          := ud_Address
                                      , us_Length           := 4
                                      );

          //no response
          if ( sd_retval <> 0 ) then
            LogError("@01F2 (SafetyBaseFSoE::ReadSDOConfig) Reading length of topology path of interface frame block failed.");
            return;
          end_if;

          // skip path length
          ud_Address += 4;

          us_BlockedTransferLength := p_SDOResponseBuffer^.ud_Data$USINT;

//*****************************************************************************
//**   TOPOLOGY PATH OF INTERFACE FRAME                                      **
//*****************************************************************************

          //send request and receive data
          sd_retval := SDOReadCfgRequ ( p_SDORequestBuffer  := p_SDORequestBuffer
                                      , p_SDOResponseBuffer := p_SDOResponseBuffer
                                      , ud_Address          := ud_Address
                                      , us_Length           := us_BlockedTransferLength
                                      , b_UseCache          := us_BlockedTransferLength < us_DataLength_Max
                                      );

          //no response
          if ( sd_retval <> 0 ) then
            LogError("@01F3 (SafetyBaseFSoE::ReadSDOConfig) Reading topology path of interface frame block failed.");
            return;
          end_if;

          // remember the destination path
          _memcpy(ptr1:=#TempPath[0], ptr2:=#p_SDOResponseBuffer^.ud_Data, cntr:=us_BlockedTransferLength);

          // skip path
          ud_Address += us_BlockedTransferLength;

//*****************************************************************************
//**   LENGTH OF COMPRESSED TOPOLOGY PATH OF INTERFACE FRAME                 **
//*****************************************************************************

          //send request and receive data
          sd_retval := SDOReadCfgRequ ( p_SDORequestBuffer  := p_SDORequestBuffer
                                      , p_SDOResponseBuffer := p_SDOResponseBuffer
                                      , ud_Address          := ud_Address
                                      , us_Length           := 4
                                      );

          //no response
          if ( sd_retval <> 0 ) then
            LogError("@01F4 (SafetyBaseFSoE::ReadSDOConfig) Reading length of compressed topology path of interface frame block failed.");
            return;
          end_if;

          // skip path length
          ud_Address += 4;

          us_BlockedTransferLength := p_SDOResponseBuffer^.ud_Data$USINT;

//*****************************************************************************
//**   COMPRESSED TOPOLOGY PATH OF INTERFACE FRAME                           **
//*****************************************************************************

          //send request and receive data
          sd_retval := SDOReadCfgRequ ( p_SDORequestBuffer  := p_SDORequestBuffer
                                      , p_SDOResponseBuffer := p_SDOResponseBuffer
                                      , ud_Address          := ud_Address
                                      , us_Length           := us_BlockedTransferLength
                                      , b_UseCache          := us_BlockedTransferLength < us_DataLength_Max
                                      );

          //no response
          if ( sd_retval <> 0 ) then
            LogError("@01F5 (SafetyBaseFSoE::ReadSDOConfig) Reading compressed topology path of interface frame block failed.");
            return;
          end_if;

          ud_Address += us_BlockedTransferLength;

          // skip max. cycle time
          ud_Address += 4;
        end_if;

        // on first 4 bytes is fix the system time
        ud_ActAddress := 4;

        // address in memory for unsafe BDINT variables
        ud_UnsafeBDINT_Offset := 0;

        // address on the module to access the fast unsafe variables via SDIAS (offset 1 for the message counter)
        ud_FastUnsafe_Offset_Out  := 1;
        ud_FastUnsafe_Offset_In   := 1;

//*****************************************************************************
//**   FSoE CONNECTION LIST                                                  **
//*****************************************************************************

        if b_IsFSoE then
          //send request and receive data
          sd_retval := SDOReadCfgRequ ( p_SDORequestBuffer  := p_SDORequestBuffer
                                      , p_SDOResponseBuffer := p_SDOResponseBuffer
                                      , ud_Address          := ud_Address
                                      , us_Length           := 4
                                      );

          //no response
          if ( sd_retval <> 0 ) then
            LogError("@0271 (SafetyBaseFSoE::ReadSDOConfig) Failed to get the number of FSoE elements.");
            return;
          end_if;

          ud_TmpCnt := p_SDOResponseBuffer^.ud_Data;

          // skip number of entries time
          ud_Address += 4;

          if ud_TmpCnt then
            for i := 1 to ud_TmpCnt do
              // read size of structure

              //send request and receive data
              sd_retval := SDOReadCfgRequ ( p_SDORequestBuffer  := p_SDORequestBuffer
                                          , p_SDOResponseBuffer := p_SDOResponseBuffer
                                          , ud_Address          := ud_Address
                                          , us_Length           := 4
                                          );

              //no response
              if ( sd_retval <> 0 ) then
                LogError("@0272 (SafetyBaseFSoE::ReadSDOConfig) Failed to read size of FSoE structure element.");
                return;
              end_if;

              // skip the whole entry since we got our info earlier via GetFSoEConnectionInfos()
              ud_Address += p_SDOResponseBuffer^.ud_Data;
            end_for;
          end_if;
        end_if;
(*

Aufbau Verbindungsliste:

Zuerst wird die Anzahl der Elemente in der Liste angegeben:

  ULONG nbrOfElements;                    // Anzahl der Elemente in der Liste

Danach kommen die einzelnen Listenelemente.
Der Anfang eines Listenelements ist auf 4 Byte ausgerichtet.

Aufbau des Listenelements:

  typedef struct FSOE_CONN_DSC
  {
    // Größe der Struktur (inkl. Längenfeld selbst)
    ULONG len;
    //! Flags
    //  Actually, type is 4 bytes in size but for compatibility reasons it is still used as 1 byte. As a result, bits 9-32 are currently not used.
    //  Bit1: 1, wenn FSoE-Master, 0=FSoE-Slave
    //  Bit2: 1, wenn die Slave-Adresse über den HW-Pfad ermittelt wird
    //  Bit3: 1, wenn CRC von der FW ermittelt werden muss
    //  Bit4: 1, wenn Interface und Slave
    //  Bit5: 1, wenn Multichannel verwendet werden, aber ein Multichannel ist nicht vorhanden und der Eingang auf 1 gesetzt wird.
    //  Bit6: 1, wenn der Adressvergabeservice verwendet werden soll
    //  Bit7: 1, wenn der Master beim Slave die Connection ID anfordert
    //  Bit8: 1, wenn es sich um ein HGW handelt
    //  Bit9: 1, wenn Assign Slave On Demand
    //  Bits 10-32: reserviert, sind auf 0 gesetzt und werden nicht ausgewertet
  #define FSOE_CONN_FLAGS_MASTER                    (1 << 0)
  #define FSOE_CONN_FLAGS_USE_HWPATH_AS_SLAVEADDR   (1 << 1)
    ULONG flags;
    //! Größe der sicheren Prozessdaten, die vom FSoE Master an den FSoE Slave übertragen werden
    // Wert kann nur 1 oder ein vielfaches von 2 sein (1, 2, 4, 6, ...)
    USHORT sizeSafeOutputs;
    //! Größe der sicheren Prozessdaten, die vom FSoE Slave an den FSoE Master übertragen werden
    // Wert kann nur 1 oder ein vielfaches von 2 sein (1, 2, 4, 6, ...)
    USHORT sizeSafeInputs;
    //! Safety over EtherCAT Slave Adresse der Safety over EtherCAT Connection
    // Bei einem Master ist das die Adresse des Ziels, bei einem Slave die eigene Adresse.
    // Wert 0 = Wert wird aus dem EEProm geholt oder über den HW-Pfad ermittelt
    // (HW-Pfad, wenn Flag FSOE_CONN_FLAGS_USE_HWPATH_AS_SLAVEADDR gesetzt ist)
    USHORT slaveAddress;

    // ==== die folgenden Daten gibt es nur im Master ====

    //! ConnectionId der Safety over EtherCAT Connection
    // Wert 0 = Wert wird aus dem EEProm geholt
    USHORT connectionId;

    //! Länge der Kommunikationsparameter, muss immer 2 sein
    USHORT commParaLength;
    //! FSoE Watchdog-Zeit in ms (nur für den Master relevant)
    USHORT watchdog_ms;
    //! Größe der Anwendungsparameter
    USHORT applParaLength;
    /*
----------------------------------------------------------------------
     * Bis hierher ist die Größe der Elemente in der Struktur fix.
     * Danach sind die Elemente mit variabler Größe angeordnet:
     *
     * Applikationsparameter:
     *    Die Applikationsparameter für ein SCP011 als FSoE Slave bestehen
     *    aus der Konfigurations-CRC (Listenheader) oder der Interface-CRC
     *    des Slaves.
     *
     * HW-Pfad: <-- ist auf 4 Byte ausgerichtet
     *    Wenn das Flag FSOE_CONN_FLAGS_USE_HWPATH_AS_SLAVEADDR gesetzt ist, dann
     *    ermittelt sich der Master die Adresse des Slaves anhand des hier
     *    angegebenen HW-Pfades.
     *    Wenn das Flag FSOE_CONN_FLAGS_USE_HWPATH_AS_SLAVEADDR nicht gesetzt ist,
     *    dann sind hier keine Daten vorhanden.
     *    Besteht aus:
     *    - normaler Pfad
     *    - komprimierter Pfad
     */

     // ==== ab hier wieder für Master und Slave ====

    /*
     * Füllbytes, damit die Größe der Struktur durch 4 teilbar ist
     */

*)

//*****************************************************************************
//**   INTERPRETER CODE                                                      **
//*****************************************************************************

        if b_IprCodeLengthAvailable = TRUE then

          sd_retval := SDOReadCfgRequ ( p_SDORequestBuffer  := p_SDORequestBuffer
                                      , p_SDOResponseBuffer := p_SDOResponseBuffer
                                      , ud_Address          := ud_Address
                                      , us_Length           := 4
                                      );

          //no response
          if ( sd_retval <> 0 ) then
            LogError("@0271 (SafetyBaseFSoE::ReadSDOConfig) Failed to get length of interpredercode.");
            return;
          end_if;

          //read length of interpretercode
          ud_TmpLength := p_SDOResponseBuffer^.ud_Data;

          //set correct address
          ud_Address += ud_TmpLength;
          ud_Address += 4;
        else

          //read til end-command is reached
          while ( 1 ) do

            //send request and receive data
            sd_retval := SDOReadCfgRequ ( p_SDORequestBuffer  := p_SDORequestBuffer
                                        , p_SDOResponseBuffer := p_SDOResponseBuffer
                                        , ud_Address          := ud_Address
                                        , us_Length           := 4
                                        );
            //no response, error
            if ( sd_retval <> 0 ) then
              LogError("@01FA (SafetyBaseFSoE::ReadSDOConfig) Reading next command failed.");
              return;
            end_if;

            //end-command found
            if ( p_SDOResponseBuffer^.ud_Data = SBF_SDO_CONFIG_END_CMD ) then
              exit;
            end_if;

            //read next opcode
            //length of one command = 4 x 4 bytes
            ud_Address += 16;

            //if there is no end-command found, the returncode of response will be <> OK, when the end of config data is missed
            //In this case the loop ends with returncode <> 0.
          end_while;

          //list of I/Os starts at last address + 16 (length of end command = 4x4 bytes)
          ud_Address += 16;

       end_if;

//*****************************************************************************
//**   LOCAL BOOL INPUTS                                                     **
//*****************************************************************************

        //read number of local bool inputs

        //send request and receive data
        sd_retval := SDOReadCfgRequ ( p_SDORequestBuffer  := p_SDORequestBuffer
                                    , p_SDOResponseBuffer := p_SDOResponseBuffer
                                    , ud_Address          := ud_Address
                                    , us_Length           := 4
                                    );

        //no response
        if ( sd_retval <> 0 ) then
          LogError("@01FB (SafetyBaseFSoE::ReadSDOConfig) Reading number of local inputs failed.");
          return;
        end_if;

        // remember the number
        BoolOuts += p_SDOResponseBuffer^.ud_Data;

        // get offset in application memory
        ud_ActAddress += p_SDOResponseBuffer^.ud_Data * 4;

        // skip number of entries
        p_SDORequestBuffer^.ud_Address += 4;

        if b_IsFSoE then
          ud_TmpCnt := p_SDOResponseBuffer^.ud_Data;

          if ud_TmpCnt then
            for i := 1 to ud_TmpCnt do
              // skip QSE, Filtertime, Modulkennung (SDIAS)
              p_SDORequestBuffer^.ud_Address += 12;

              //send request and receive data
              sd_retval := SDOReadCfgRequ ( p_SDORequestBuffer  := p_SDORequestBuffer
                                          , p_SDOResponseBuffer := p_SDOResponseBuffer
                                          , ud_Address          := p_SDORequestBuffer^.ud_Address
                                          , us_Length           := 4
                                          );

              //no response
              if ( sd_retval <> 0 ) then
                LogError("@0273 (SafetyBaseFSoE::ReadSDOConfig) Reading number of FSoE connections for local inputs failed.");
                return;
              end_if;

              // skip number of entries and the entries
              p_SDORequestBuffer^.ud_Address += 4 + 4 * p_SDOResponseBuffer^.ud_Data;
            end_for;
          end_if;
        else
          // only available at new modules
          if b_CfgTypeV2 then
            ud_skipLength := 12 * p_SDOResponseBuffer^.ud_Data; // QSE, Filtertime, Modulkennung(SDIAS)
          else
            ud_skipLength := 8 * p_SDOResponseBuffer^.ud_Data; // QSE, Filtertime
          end_if;

          p_SDORequestBuffer^.ud_Address += ud_skipLength;
        end_if;

//*****************************************************************************
//**   LOCAL BOOL OUTPUTS AS INPUTS                                          **
//*****************************************************************************

        // get number of safe outputs as inputs

        //send request and receive data
        sd_retval := SDOReadCfgRequ ( p_SDORequestBuffer  := p_SDORequestBuffer
                                    , p_SDOResponseBuffer := p_SDOResponseBuffer
                                    , ud_Address          := p_SDORequestBuffer^.ud_Address
                                    , us_Length           := 4
                                    );

        //no response
        if ( sd_retval <> 0 ) then
          LogError("@01FC (SafetyBaseFSoE::ReadSDOConfig) Reading number of safe outputs as inputs failed.");
          return;
        end_if;

        // remember the number
        BoolOuts += p_SDOResponseBuffer^.ud_Data;

        // get offset in application memory
        ud_ActAddress += p_SDOResponseBuffer^.ud_Data * 4;

        p_SDORequestBuffer^.ud_Address += 4;

        if b_IsFSoE then
          ud_TmpCnt := p_SDOResponseBuffer^.ud_Data;

          if ud_TmpCnt then
            for i := 1 to ud_TmpCnt do
              //send request and receive data
              sd_retval := SDOReadCfgRequ ( p_SDORequestBuffer  := p_SDORequestBuffer
                                          , p_SDOResponseBuffer := p_SDOResponseBuffer
                                          , ud_Address          := p_SDORequestBuffer^.ud_Address
                                          , us_Length           := 4
                                          );

              //no response
              if ( sd_retval <> 0 ) then
                LogError("@0274 (SafetyBaseFSoE::ReadSDOConfig) Reading number of FSoE connections for local outputs as inputs failed.");
                return;
              end_if;

              // skip number of entries and the entries
              p_SDORequestBuffer^.ud_Address += 4 + 4 * p_SDOResponseBuffer^.ud_Data;
            end_for;
          end_if;
        end_if;

//*****************************************************************************
//**   SAFE BOOL OUTPUT VARIABLES                                            **
//*****************************************************************************

        // get number of safe bool output vars

        //send request and receive data
        sd_retval := SDOReadCfgRequ ( p_SDORequestBuffer  := p_SDORequestBuffer
                                    , p_SDOResponseBuffer := p_SDOResponseBuffer
                                    , ud_Address          := p_SDORequestBuffer^.ud_Address
                                    , us_Length           := 4
                                    );

        //no response
        if ( sd_retval <> 0 ) then
          LogError("@01FD (SafetyBaseFSoE::ReadSDOConfig) Reading number of safe bool output vars failed.");
          return;
        end_if;

        // remember the number
        BoolOuts += p_SDOResponseBuffer^.ud_Data;

        // get offset in application memory
        ud_ActAddress += p_SDOResponseBuffer^.ud_Data * 4;

        p_SDORequestBuffer^.ud_Address += 4;

        if b_IsFSoE then
          ud_TmpCnt := p_SDOResponseBuffer^.ud_Data;

          if ud_TmpCnt then
            for i := 1 to ud_TmpCnt do
              //send request and receive data
              sd_retval := SDOReadCfgRequ ( p_SDORequestBuffer  := p_SDORequestBuffer
                                          , p_SDOResponseBuffer := p_SDOResponseBuffer
                                          , ud_Address          := p_SDORequestBuffer^.ud_Address
                                          , us_Length           := 4
                                          );

              //no response
              if ( sd_retval <> 0 ) then
                LogError("@0275 (SafetyBaseFSoE::ReadSDOConfig) Reading number of FSoE connections for bool outputs failed.");
                return;
              end_if;

              // skip number of entries and the entries
              p_SDORequestBuffer^.ud_Address += 4 + 4 * p_SDOResponseBuffer^.ud_Data;
            end_for;
          end_if;
        end_if;

        // the new container has some additional content here
        if b_CfgTypeV3 then

//*****************************************************************************
//**   LOCAL DINT INPUTS                                                     **
//*****************************************************************************

          //read number of local dint inputs

          //send request and receive data
          sd_retval := SDOReadCfgRequ ( p_SDORequestBuffer  := p_SDORequestBuffer
                                      , p_SDOResponseBuffer := p_SDOResponseBuffer
                                      , ud_Address          := p_SDORequestBuffer^.ud_Address
                                      , us_Length           := 4
                                      );

          //no response
          if ( sd_retval <> 0 ) then
            LogError("@01FE (SafetyBaseFSoE::ReadSDOConfig) Reading number of local DINT inputs failed.");
            return;
          end_if;

          // remember the number
          DintOuts += p_SDOResponseBuffer^.ud_Data;

          // get offset in application memory
          ud_ActAddress += p_SDOResponseBuffer^.ud_Data * 8;

          p_SDORequestBuffer^.ud_Address += 4;

          if b_IsFSoE then
            ud_TmpCnt := p_SDOResponseBuffer^.ud_Data;

            if ud_TmpCnt then
              for i := 1 to ud_TmpCnt do
                // skip QSE, Filtertime, Modulkennung (SDIAS)
                p_SDORequestBuffer^.ud_Address += 12;

                //send request and receive data
                sd_retval := SDOReadCfgRequ ( p_SDORequestBuffer  := p_SDORequestBuffer
                                            , p_SDOResponseBuffer := p_SDOResponseBuffer
                                            , ud_Address          := p_SDORequestBuffer^.ud_Address
                                            , us_Length           := 4
                                            );

                //no response
                if ( sd_retval <> 0 ) then
                  LogError("@0276 (SafetyBaseFSoE::ReadSDOConfig) Reading number of FSoE connections for local DINT inputs failed.");
                  return;
                end_if;

                // skip number of entries and the entries
                p_SDORequestBuffer^.ud_Address += 4 + 4 * p_SDOResponseBuffer^.ud_Data;
              end_for;
            end_if;
          else
            p_SDORequestBuffer^.ud_Address += 12 * p_SDOResponseBuffer^.ud_Data;
          end_if;

//*****************************************************************************
//**   LOCAL DINT OUTPUTS AS INPUTS                                          **
//*****************************************************************************

          // get number of safe dint outputs as inputs

          //send request and receive data
          sd_retval := SDOReadCfgRequ ( p_SDORequestBuffer  := p_SDORequestBuffer
                                      , p_SDOResponseBuffer := p_SDOResponseBuffer
                                      , ud_Address          := p_SDORequestBuffer^.ud_Address
                                      , us_Length           := 4
                                      );

          //no response
          if ( sd_retval <> 0 ) then
            LogError("@01FF (SafetyBaseFSoE::ReadSDOConfig) Reading number of safe DINT outputs as inputs failed.");
            return;
          end_if;

          // remember the number
          DintOuts += p_SDOResponseBuffer^.ud_Data;

          // get offset in application memory
          ud_ActAddress += p_SDOResponseBuffer^.ud_Data * 8;

          p_SDORequestBuffer^.ud_Address += 4;

          if b_IsFSoE then
            ud_TmpCnt := p_SDOResponseBuffer^.ud_Data;

            if ud_TmpCnt then
              for i := 1 to ud_TmpCnt do
                //send request and receive data
                sd_retval := SDOReadCfgRequ ( p_SDORequestBuffer  := p_SDORequestBuffer
                                            , p_SDOResponseBuffer := p_SDOResponseBuffer
                                            , ud_Address          := p_SDORequestBuffer^.ud_Address
                                            , us_Length           := 4
                                            );

                //no response
                if ( sd_retval <> 0 ) then
                  LogError("@0277 (SafetyBaseFSoE::ReadSDOConfig) Reading number of FSoE connections for local DINT outputs as inputs failed.");
                  return;
                end_if;

                // skip number of entries and the entries
                p_SDORequestBuffer^.ud_Address += 4 + 4 * p_SDOResponseBuffer^.ud_Data;
              end_for;
            end_if;
          end_if;

        end_if;

//*****************************************************************************
//**   SAFE DINT OUTPUT VARIABLES                                            **
//*****************************************************************************

        // get number of safe dint output vars

        //send request and receive data
        sd_retval := SDOReadCfgRequ ( p_SDORequestBuffer  := p_SDORequestBuffer
                                    , p_SDOResponseBuffer := p_SDOResponseBuffer
                                    , ud_Address          := p_SDORequestBuffer^.ud_Address
                                    , us_Length           := 4
                                    );

        //no response
        if ( sd_retval <> 0 ) then
          LogError("@0200 (SafetyBaseFSoE::ReadSDOConfig) Reading number of safe dint output vars failed.");
          return;
        end_if;

        // only when there is a manager
        if pSafetyManagerThis then
          // remember the number
          DintOuts += p_SDOResponseBuffer^.ud_Data;

          // now we're ready to determine the PDO size of this module
          TempModuleConfig.PdoOutLen := CalcPDOLength(BoolOuts, DintOuts);

          // if it's our own path, remember the PDO length
//          if (PathOfThisCPU[0]$UINT = (pListHeader^.p_us_Path$^UINT)^) & (ToStdLib.MemCmp(#PathOfThisCPU[0], pListHeader^.p_us_Path, PathOfThisCPU[0]$UINT + 2) = 0) then
//            MyPDOReadSize := TempModuleConfig.PdoOutLen;
//          end_if;
        end_if;

        // get offset in application memory
        ud_ActAddress += p_SDOResponseBuffer^.ud_Data * 8;

        p_SDORequestBuffer^.ud_Address += 4;

        if b_IsFSoE then
          ud_TmpCnt := p_SDOResponseBuffer^.ud_Data;

          if ud_TmpCnt then
            for i := 1 to ud_TmpCnt do
              //send request and receive data
              sd_retval := SDOReadCfgRequ ( p_SDORequestBuffer  := p_SDORequestBuffer
                                          , p_SDOResponseBuffer := p_SDOResponseBuffer
                                          , ud_Address          := p_SDORequestBuffer^.ud_Address
                                          , us_Length           := 4
                                          );

              //no response
              if ( sd_retval <> 0 ) then
                LogError("@0278 (SafetyBaseFSoE::ReadSDOConfig) Reading number of FSoE connections for DINT outputs failed.");
                return;
              end_if;

              // skip number of entries and the entries
              p_SDORequestBuffer^.ud_Address += 4 + 4 * p_SDOResponseBuffer^.ud_Data;
            end_for;
          end_if;
        end_if;

        ud_Address := p_SDORequestBuffer^.ud_Address;

        // special unsafe variables (not supported by old modules)
        if b_CfgTypeV2 then

//*****************************************************************************
//**   FAST UNSAFE OUTPUT VARIABLES                                          **
//*****************************************************************************
          //check if used a SCP111 or SCP211
          if b_IprCodeLengthAvailable = FALSE then
            // get number of fast unsafe output vars

            //send request and receive data
            sd_retval := SDOReadCfgRequ ( p_SDORequestBuffer  := p_SDORequestBuffer
                                        , p_SDOResponseBuffer := p_SDOResponseBuffer
                                        , ud_Address          := ud_Address
                                        , us_Length           := 4
                                        );

            //no response
            if ( sd_retval <> 0 ) then
              LogError("@0201 (SafetyBaseFSoE::ReadSDOConfig) Reading number of fast unsafe output vars failed.");
              return;
            end_if;

            // get offset in application memory
            ud_ActAddress += p_SDOResponseBuffer^.ud_Data * 4;

            // if it's our own path, remember the fast unsafe settings
            if (PathOfThisCPU[0]$UINT = (pListHeader^.p_us_Path$^UINT)^) & (ToStdLib.MemCmp(#PathOfThisCPU[0], pListHeader^.p_us_Path, PathOfThisCPU[0]$UINT + 2) = 0) then
              if (p_SDOResponseBuffer^.ud_Data <> 0) then
                if ActivateFastUnsafeIOs then
                  b_FastUnsafeOutputsActive := TRUE;
                else
                  // error => can't go on like this
                  LogError("@0202 (SafetyBaseFSoE::ReadSDOConfig) Number or size of module accesses increased with new safety project!");
                  LogError("@0203 (SafetyBaseFSoE::ReadSDOConfig) => Can't continue, because the new data is not covered by the actual accesses! Restart Application!");

                  b_NeedApplicationRestart := TRUE;
                end_if;
              end_if;
            end_if;

            ud_Address += 4;

          else

//*****************************************************************************
//**   FAST UNSAFE BOOL OUTPUT VARIABLES  SCP211                             **
//*****************************************************************************
            //read number of unsafe output vars

            //send request and receive data
            sd_retval := SDOReadCfgRequ ( p_SDORequestBuffer  := p_SDORequestBuffer
                                        , p_SDOResponseBuffer := p_SDOResponseBuffer
                                        , ud_Address          := ud_Address
                                        , us_Length           := 4
                                        );

            //no response
            if ( sd_retval <> 0 ) then
              LogError("@0204 (SafetyBaseFSoE::ReadSDOConfig) Reading number of unsafe bool output vars failed.");
              return;
            end_if;

            ud_CntFastUnsafeOutputs := p_SDOResponseBuffer^.ud_Data;

            ud_Address += 4;

            // skip the names of unsafe outputs
            for i := 1 to ud_CntFastUnsafeOutputs do

              // get length of Name
              sd_retval := SDOReadCfgRequ ( p_SDORequestBuffer  := p_SDORequestBuffer
                                          , p_SDOResponseBuffer := p_SDOResponseBuffer
                                          , ud_Address          := ud_Address
                                          , us_Length           := 4
                                          );
              //no response
              if ( sd_retval <> 0 ) then
                LogError("@0205 (SafetyBaseFSoE::ReadSDOConfig) Reading length of unsafe bool output name failed.");
                return;
              end_if;

              // prepare address to get name
              ud_Address += 4;

    //          ud_ActStrLen := ud_TmpStrLen := p_SDOResponseBuffer^.ud_Data;
              ud_TmpStrLen := p_SDOResponseBuffer^.ud_Data;
              ud_ActStrLen := ud_TmpStrLen;
              ud_TmpAddress := ud_Address;

              IF p_BlockedTransferMemory = NIL THEN
                sd_retval := -100;
                SetSafetyState(NewState:=_MemAllocFailed);
                RETURN;
              END_IF;

              IF ud_BlockedTransferMemorySize < (ud_TmpStrLen + 1) THEN
                p_BlockedTransferMemory := ToStdLib.ReAlloc(mptr:=p_BlockedTransferMemory, newsize:=GetNewMemSize(ud_TmpStrLen + 1));
                IF p_BlockedTransferMemory = NIL THEN
                  ud_BlockedTransferMemorySize := 0;
                  sd_retval := -100;
                  SetSafetyState(NewState:=_MemAllocFailed);
                  RETURN;
                ELSE
                  ud_BlockedTransferMemorySize := GetNewMemSize(ud_TmpStrLen + 1);
                END_IF;
              END_IF;

              ToStdLib.MemSet(dest:=p_BlockedTransferMemory, value:=0, size:=ud_BlockedTransferMemorySize);

              p_TmpBlockedData := p_BlockedTransferMemory;

              us_BlockedTransferLength := BlockedTransferLength(ud_Datalength:=ud_TmpStrLen, us_MaxBlocklength:=60);

              while us_BlockedTransferLength do

                // get name
                sd_retval := SDOReadCfgRequ ( p_SDORequestBuffer  := p_SDORequestBuffer
                                            , p_SDOResponseBuffer := p_SDOResponseBuffer
                                            , ud_Address          := ud_TmpAddress
                                            , us_Length           := us_BlockedTransferLength
                                            , b_UseCache          := us_BlockedTransferLength < us_DataLength_Max
                                            );
                //no response
                if ( sd_retval <> 0 ) then
                  LogError("0206 (SafetyBaseFSoE::ReadSDOConfig) Reading unsafe bool output name failed.");
                  return;
                end_if;

                ToStdLib.MemCpy(dest:=p_TmpBlockedData,
                                 source:=#p_SDOResponseBuffer^.ud_Data,
                                 size:=us_BlockedTransferLength);

                p_TmpBlockedData += us_BlockedTransferLength;
                ud_TmpAddress += us_BlockedTransferLength;
                ud_TmpStrLen -= us_BlockedTransferLength;

                us_BlockedTransferLength := BlockedTransferLength(ud_Datalength:=ud_TmpStrLen, us_MaxBlocklength:=60);

              end_while;

              sd_retval :=AddFastUnsafeRoutElement(pRoutTable:=#p_FastUnsafeOutputsTable,
                                                   pRoutElementsNo:=#ui_CntFastUnsafeOutputs,
                                                   ud_Address:=ud_FastUnsafe_Offset_Out,
                                                   ui_NameLen:=ud_ActStrLen$UINT,
                                                   pNameNewElement:=p_BlockedTransferMemory$^CHAR,
                                                   bWriteVar:=TRUE);

              // if unsafe component not found (sd_retval <> 0), it's not problem for whole safe application

              // get offset in application memory
              ud_ActAddress += 4;
              ud_FastUnsafe_Offset_Out += 4;

              // prepare address for next unsafe output or for number of safe inputs
              ud_Address += ud_ActStrLen;

            end_for;

  //*****************************************************************************
  //**   FAST UNSAFE BDINT OUTPUT VARIABLES   SCP211                           **
  //*****************************************************************************

            //read number of unsafe BDINT output vars

            //send request and receive data
            sd_retval := SDOReadCfgRequ ( p_SDORequestBuffer  := p_SDORequestBuffer
                                        , p_SDOResponseBuffer := p_SDOResponseBuffer
                                        , ud_Address          := ud_Address
                                        , us_Length           := 4
                                        );

            //no response
            if ( sd_retval <> 0 ) then
              LogError("@0207 (SafetyBaseFSoE::ReadSDOConfig) Reading number of unsafe BDINT output vars failed.");
              return;
            end_if;

            ud_CntFastUnsafeOutputs := p_SDOResponseBuffer^.ud_Data;

            ud_Address += 4;

            if ud_CntFastUnsafeOutputs then

              //SDO request for this command has 5 bytes additional data
              pBitMasks$^void := ToStdLib.Malloc(size := ud_CntFastUnsafeOutputs * sizeof(BDINT));

              if ( pBitMasks = NIL ) then
                sd_retval                         := -100;
                SetSafetyState(NewState:=_MemAllocFailed);
                LogError("@0208 (SafetyBaseFSoE::ReadSDOConfig) Failed to allocate memory for the BDINT variable bitmasks.");
                return;
              end_if;

              // get the bitmasks for the BDINT variables
              for i := 1 to ud_CntFastUnsafeOutputs do

                // get bitmask
                sd_retval := SDOReadCfgRequ ( p_SDORequestBuffer  := p_SDORequestBuffer
                                            , p_SDOResponseBuffer := p_SDOResponseBuffer
                                            , ud_Address          := ud_Address
                                            , us_Length           := 4
                                            );
                //no response
                if ( sd_retval <> 0 ) then
                  LogError("@0207 (SafetyBaseFSoE::ReadSDOConfig) Reading bit mask of unsafe BDINT output failed.");
                  return;
                end_if;

                // prepare address for the next one
                ud_Address += 4;

                // save the bitmask for adding the rout element
                (pBitMasks + (i-1) * sizeof(BDINT))^ := p_SDOResponseBuffer^.ud_Data;
              end_for;

              // skip the names of unsafe outputs
              for i := 1 to ud_CntFastUnsafeOutputs do
